FUNCTION_BLOCK FB_UDPTxStateMachine
VAR_IN_OUT
	fbTxFIFO		: FB_UDPFrameFIFO;
END_VAR
VAR_INPUT
	bEnable			: BOOL			:= FALSE;			// TRUE => Enable/connect, FALSE => Disable/disconnect
	tReconnect		: TIME			:= T#5S;			// Reconnect delay time
	bLog			: BOOL			:= FALSE;			// TRUE => Enable log message output, FALSE => Disable 
	sPrefix			: STRING 		:= 'PeerToPeerX::'; // Log message description string (allows the identification of log message source)
END_VAR
VAR_OUTPUT
	bCreated		: BOOL;		// Connectionless socket state (TRUE => created, FALSE => closed)
END_VAR
VAR
	fbCreate		: FB_SocketUdpCreate;
	hSocket			: T_HSOCKET;
	fbClose			: FB_SocketClose;
	fbSendTo		: FB_SocketUdpSendTo;
	stSendTo		: ST_UDPFrameEntry;
	fbCreateTimer	: TON := ( PT := T#0S );	
	eState			: E_UDPClientServerState;
END_VAR

CASE eState OF
	(* Idle State *)
	eUDP_STATE_IDLE:
		IF bEnable XOR bCreated THEN
			IF bEnable THEN
				(* Clear send fifo *)
				fbTxFIFO.Clear( sPrefix := CONCAT( sPrefix, 'FB_FrameFifo(sender)::' ), bLog := bLog );
				
				(* At program start (first time) connect immediately, next time after delay time *)
				fbCreateTimer( IN := TRUE );
				IF fbCreateTimer.Q THEN
					fbCreateTimer( IN := FALSE, PT := tReconnect ); 
					eState := eUDP_STATE_CREATE_START;
				END_IF
			ELSE
				eState := eUDP_STATE_CLOSE_START;
			END_IF
		ELSIF bCreated THEN
			fbTxFIFO.RemoveHead( stGet => stSendTo );
			IF fbTxFIFO.bOk THEN
				eState := eUDP_STATE_SEND_START;
			END_IF
		ELSE
			fbCreateTimer( IN := FALSE, PT := T#0S );
		END_IF
	
	(* Creation States *)
	eUDP_STATE_CREATE_START:
		fbCreate( bExecute := FALSE  );
		fbCreate( sSrvNetId := sSrvNetId, sLocalHost:= sLocalHost, nLocalPort:= nLocalTxPort, bExecute:= TRUE );
		eState := eUDP_STATE_CREATE_WAIT;

	eUDP_STATE_CREATE_WAIT:
		fbCreate( bExecute := FALSE );
		IF NOT fbCreate.bBusy THEN
			IF NOT fbCreate.bError THEN
				bCreated := TRUE;
				hSocket := fbCreate.hSocket;
// 				fbLog.Message( sMessage := 'Connectionless (UDP) socket created!', hSocket := fbCreate.hSocket );
				eState := eUDP_STATE_IDLE;
			ELSE
// 				fbLog.Error( sMessage := 'FB_SocketUdpCreate()', nErrID := fbCreate.nErrID );
				eState := eUDP_STATE_ERROR;
			END_IF
		END_IF
	
	(* Sending States *)
	eUDP_STATE_SEND_START:
		fbSendTo( bExecute := FALSE );
		fbSendTo( sSrvNetId := sSrvNetId, sRemoteHost := stSendTo.stRemoteAddr.sAddr,
					nRemotePort := stSendTo.stRemoteAddr.nPort,
					pSrc:= ADR( stSendTo.sMessage ),
					//cbLen:= INT_TO_UDINT(LEN( stSendTo.sMessage )) + 1, (* Include the end delimiter *)
					cbLen := SIZEOF(UDP_DATA),
					hSocket:= fbCreate.hSocket, bExecute:= TRUE );
		eState := eUDP_STATE_SEND_WAIT;

	eUDP_STATE_SEND_WAIT:
		fbSendTo( bExecute := FALSE );
		IF NOT fbSendTo.bBusy THEN
			IF NOT fbSendTo.bError THEN
				eState := eUDP_STATE_IDLE;
			ELSE
// 				fbLog.Error( sMessage := 'FB_SocketUdpSendTo()', nErrID := fbSendTo.nErrID );
				eState := eUDP_STATE_ERROR;
			END_IF
		END_IF
		
	(* Closing States *)
	eUDP_STATE_CLOSE_START:
// 		fbLog.Message( sMessage := 'Closing connectionless (UDP) socket!', hSocket := fbCreate.hSocket );
		fbClose( bExecute := FALSE );
		fbClose( sSrvNetId := sSrvNetId, hSocket := fbCreate.hSocket, bExecute := TRUE );
		eState := eUDP_STATE_CLOSE_WAIT;
		
	eUDP_STATE_CLOSE_WAIT:
		fbClose( bExecute := FALSE );
		IF NOT fbClose.bBusy THEN
			bCreated := FALSE;
			IF NOT fbClose.bError THEN
				eState := eUDP_STATE_IDLE;
			ELSE
// 				fbLog.Error( sMessage := 'FB_SocketClose()', nErrID := fbClose.nErrID );
				eState := eUDP_STATE_ERROR;
			END_IF
		END_IF

	(* Error State *)

	eUDP_STATE_ERROR: (* Error step *)
		IF bCreated THEN
			eState := eUDP_STATE_CLOSE_START;
		ELSE
			eState := eUDP_STATE_IDLE;
		END_IF

END_CASE

//FB_Exit must be implemented explicitly. If there is an implementation, then the
//method is called before the controller removes the code of the function block instance
//(implicit call). The return value is not evaluated.
METHOD FB_Exit: BOOL
VAR_INPUT
    bInCopyCode: BOOL;  // TRUE: the exit method is called in order to leave the instance which will be copied afterwards (online change).  
END_VAR
IF bCreated THEN
    fbClose(sSrvNetId := '', hSocket := hSocket, bExecute := TRUE);
END_IF
END_METHOD

//FB_Init is always available implicitly and it is used primarily for initialization.
//The return value is not evaluated. For a specific influence, you can also declare the
//methods explicitly and provide additional code there with the standard initialization
//code. You can evaluate the return value.
METHOD FB_Init: BOOL
VAR_INPUT
    bInitRetains: BOOL; // TRUE: the retain variables are initialized (reset warm / reset cold)
    bInCopyCode: BOOL;  // TRUE: the instance will be copied to the copy code afterward (online change)   
END_VAR
END_METHOD

END_FUNCTION_BLOCK

(* stored: Version 1.1.0.1
   POU FB_UDPTxStateMachine: Id {eaa388e7-d7d6-421e-b48b-746a67ef0c5a}, SpecialFunc None
   Method FB_Exit: Id {08b2b0a0-5425-4e13-b9eb-61b7cc809be2}
   Method FB_Init: Id {2252a51d-108b-45e9-8470-ed4d45193779} *)
